// TIA Portal V19 export
DATA_BLOCK "HS_SKIDS"   // DB23
{ S7_Optimized_Access := 'FALSE' }
   VAR RETAIN
      HS_SKIDS : Struct
         TEMP_SP : Real := 120.0;
         START : Bool;
         RUNNING : Bool;
         EMG : Bool;
         HOLD_RESUME : Bool;
         RUUNING : Bool;
         PUMP_SEL : Int;
         AUTO : Bool;
         HEADER_PSP : Real := 2.5;
         START_PLS : Bool;
         STOP_PLS : Bool;
         "PUMP 1 RPM" : Real;
         "PUMP 1RPM_SP" : Real := 49.9;
         "PUMP 2 RPM" : Real;
         "PUMP 2 RPM_SP" : Real := 49.9;
         "PUMP 3 RPM" : Real;
         "PUMP 3 RPM_SP" : Real := 49.9;
         CV_CMD : Bool;
         RESET : Bool;
      END_STRUCT;
   END_VAR
BEGIN
END_DATA_BLOCK
